Fanuc KAREL source: compact_preamble.KL

PROGRAM KB00202
%NOLOCKGROUP
VAR
P1 : FILE
P2 : STRING[80]
P3 : STRING[80]
P4:INTEGER
BEGIN
P2='A'
P3='A'
P4=1
XML_SETVAR(P1,P2,P3,P4)
END KB00202
